(* IEC 61131-3 sources: plc-iiot-stack/tests/POUs/FB_JsonFlatParser_Test, 13 files *)

(* ---- AcceptsWhitespaceAndEmptyObject.method.decl.st ---- *)
// Пробелы, табуляции и переводы строк между токенами; пустой объект.
METHOD PRIVATE AcceptsWhitespaceAndEmptyObject
VAR_INST
    fbParser : FB_JsonFlatParser;
    sJsonIn : STRING(GVL_Const.MQTT_CMD_PAYLOAD_LEN);
END_VAR

(* ---- DecodesEscapes.method.decl.st ---- *)
// Escape-последовательности JSON; код вне ASCII и неизвестные — BadEscape.
METHOD PRIVATE DecodesEscapes
VAR_INST
    fbParser : FB_JsonFlatParser;
    sJsonIn : STRING(GVL_Const.MQTT_CMD_PAYLOAD_LEN);
END_VAR
VAR
    sText : STRING(GVL_Const.JSON_STR_LEN);
END_VAR

(* ---- FailedParseClearsPreviousFields.method.decl.st ---- *)
// После неудачного разбора поля прошлого объекта не видны.
METHOD PRIVATE FailedParseClearsPreviousFields
VAR_INST
    fbParser : FB_JsonFlatParser;
    sJsonIn : STRING(GVL_Const.MQTT_CMD_PAYLOAD_LEN);
END_VAR

(* ---- LimitsFieldCount.method.decl.st ---- *)
// Полей не больше 12; 13-е — TooManyFields.
METHOD PRIVATE LimitsFieldCount
VAR_INST
    fbParser : FB_JsonFlatParser;
    sJsonIn : STRING(GVL_Const.MQTT_CMD_PAYLOAD_LEN);
END_VAR

(* ---- LimitsKeyAndValueLength.method.decl.st ---- *)
// Ключ до 31 и строка до 64 символов; длиннее — KeyTooLong, ValueTooLong.
METHOD PRIVATE LimitsKeyAndValueLength
VAR_INST
    fbParser : FB_JsonFlatParser;
    sJsonIn : STRING(GVL_Const.MQTT_CMD_PAYLOAD_LEN);
END_VAR

(* ---- ParsesFlatObjectWithAllTypes.method.decl.st ---- *)
// Строка, число с порядком, true, false, null; поиск по ключу, ключ по номеру.
METHOD PRIVATE ParsesFlatObjectWithAllTypes
VAR_INST
    fbParser : FB_JsonFlatParser;
    sJsonIn : STRING(GVL_Const.MQTT_CMD_PAYLOAD_LEN);
END_VAR
VAR
    sText : STRING(GVL_Const.JSON_STR_LEN);
    lrNum : LREAL;
    xFlag : BOOL;
END_VAR

(* ---- RejectsDuplicateKeys.method.decl.st ---- *)
// Повторяющийся ключ — Duplicate (неоднозначная команда).
METHOD PRIVATE RejectsDuplicateKeys
VAR_INST
    fbParser : FB_JsonFlatParser;
    sJsonIn : STRING(GVL_Const.MQTT_CMD_PAYLOAD_LEN);
END_VAR

(* ---- RejectsNestedObjectsAndArrays.method.decl.st ---- *)
// Вложенный объект и массив — Nested.
METHOD PRIVATE RejectsNestedObjectsAndArrays
VAR_INST
    fbParser : FB_JsonFlatParser;
    sJsonIn : STRING(GVL_Const.MQTT_CMD_PAYLOAD_LEN);
END_VAR

(* ---- RejectsRawControlCharacters.method.decl.st ---- *)
// Управляющий символ внутри строки без экранирования — Syntax.
METHOD PRIVATE RejectsRawControlCharacters
VAR_INST
    fbParser : FB_JsonFlatParser;
    sJsonIn : STRING(GVL_Const.MQTT_CMD_PAYLOAD_LEN);
END_VAR

(* ---- RejectsSyntaxErrors.method.decl.st ---- *)
// Пустой вход, не объект, незакрытый объект, нет двоеточия, лишняя запятая, ключ без кавычек.
METHOD PRIVATE RejectsSyntaxErrors
VAR_INST
    fbParser : FB_JsonFlatParser;
    sJsonIn : STRING(GVL_Const.MQTT_CMD_PAYLOAD_LEN);
END_VAR

(* ---- RejectsTrailingCharacters.method.decl.st ---- *)
// Символы после объекта — Trailing с позицией.
METHOD PRIVATE RejectsTrailingCharacters
VAR_INST
    fbParser : FB_JsonFlatParser;
    sJsonIn : STRING(GVL_Const.MQTT_CMD_PAYLOAD_LEN);
END_VAR

(* ---- TracksIntegerLiterals.method.decl.st ---- *)
// Целое JSON — без дробной части и порядка: 1792137621000 — да, 1.0 и 1e3 — нет.
METHOD PRIVATE TracksIntegerLiterals
VAR_INST
    fbParser : FB_JsonFlatParser;
    sJsonIn : STRING(GVL_Const.MQTT_CMD_PAYLOAD_LEN);
END_VAR
VAR
    lrNum : LREAL;
END_VAR

(* ---- ValidatesNumberGrammarAndRange.method.decl.st ---- *)
// Числа: ведущий ноль, точка без цифр, знак без цифр, порядок без цифр, вне REAL, много цифр.
METHOD PRIVATE ValidatesNumberGrammarAndRange
VAR_INST
    fbParser : FB_JsonFlatParser;
    sJsonIn : STRING(GVL_Const.MQTT_CMD_PAYLOAD_LEN);
END_VAR
VAR
    lrNum : LREAL;
END_VAR
